(* IEC 61131-3 sources: NachHouse_TST/ExamplesCustomLogin/CustomLogin, 2 files *)

(* ---- CustomLogin.st ---- *)
VAR_GLOBAL
  CustomizedLoginPage AT %S355.1 : BOOL := true;
END_VAR

VAR_GLOBAL RETAIN
   myName  : STRING[10] := 'Service';
   myPass  : STRING[10] := 'service';
END_VAR

VAR_GLOBAL
  passSet : BOOL;
  passCancel : BOOL;
  webName : STRING[10];
  webPass : STRING[10];
END_VAR

(* ---- prgMain.ST ---- *)
PROGRAM prgMain
  VAR
  END_VAR

  IF passCancel THEN
    webName := myName;
    webPass := '';
    passCancel := false;
  END_IF;

  IF NOT passSet THEN
    IF LEN(webName) > 0 AND LEN(webPass) > 0 THEN //if set from web, copy values to retain
      myName := webName;
      myPass := webPass;
    END_IF;
    SetWebPSW(user := 0, name := myName, password := myPass);
    webName := myName;
    webPass := '';
    passSet := true;
  END_IF;

END_PROGRAM
